Staubli VAL3: appLauncher.pjx

--- appLauncher.pjx ---
Parameters version=s8.21Cs9_BS4703 stackSize=200000 millimeterUnit=true
Program file=_getForce.pgx
Program file=_productCycle.pgx
Program file=_supervisorTasks.pgx
Program file=_systemStates.pgx
Program file=_tCycleCtrl.pgx
Program file=_TolleranceCheck.pgx
Program file=Init.pgx
Program file=kill.pgx
Program file=Main.pgx
Program file=search_traj.pgx
Program file=start.pgx
Program file=stop.pgx
Data file=appLauncher.dtx
Library alias=rs path=Disk://source/projectSource/robotStatus/robotStatus.pjx
Library alias=io path=Disk://source/projectSource/io/io.pjx
Library alias=home path=Disk://HMI_cs9/home/home.pjx
Library alias=plc path=Disk://source/projectSource/plc/plc.pjx
Library alias=prog path=Disk://source/projectSource/program/program.pjx
Library alias=program path=Disk://source/projectSource/program/program.pjx
Library alias=hmi_util path=Disk://HMI_cs9/HMI_util/HMI_util.pjx
Library alias=libTqe path=Disk://LibTorque/LibTorque.pjx
Library alias=trajectory path=Disk://source/projectSource/trajectory/trajectory.pjx
Library alias=ar path=Disk://autoReturn/autoReturn.pjx
Library alias=saveData path=Disk://source/saveData/saveData.pjx

--- appLauncher.dtx ---
bool _bAtHome
bool _bEndCycle
bool _bHeavyAlarm
bool _bIsScara
bool _bShowEndBt
bool _bShowPauseBt
bool _bShowResetBt
bool _bShowStartBt
bool _bShowStopBt
bool bBool
bool bControlByRobot = true
bool bTosave
frame test3 = {fatherId=world[0]}
num _nAvgCapacity
num _nBestCapacity
num _nCTIndex
num _nCapacity
num _nClock[10]
  [1] = 12488.271809
  [3] = 12488.271821
num _nCycleTime[10]
num _nLastStateCMD
num _nOmacStat
num _nStateCMD
num nCycleCmd
num nErrorCode = 1
num nLastLib
num nProgCode
string _sArmType
string _sOmacCmd
string _sOmacStatus = "1"
string _sPageAvergeCapacity
string _sPageBestCapacity
string _sPageCurrentCapacity
string _sPageCycleStatus
string _sPageHerej
string _sPagePosition
string _sPageProfile
string _sPageRobotStatus
string _sPageSN
string sMsg
num nForce[6]
public bool bGetMovId
mdesc mHome = {accel=20, vel=20, decel=20, blend=off}
string sSessionList
pointRx pPowerOFF = {fatherId=world[0]}
bool bMemState
pointRx pHere1 = {fatherId=world[0]}
pointRx pHere2 = {fatherId=world[0]}
bool bAutoConnectMove

--- Main.pgx ---
program Main()
  local bool l_bResult
  local bool l_bStartClock
  local num l_nClock
  local num l_nResult
begin
  //

  home:sVersion="version:5.0"
  resetMotion()
  //初始化
  //  call cycle_Init()
  //
  // userPage("StartUp")

  sMsg=">>> Loading 数据库 "+toString("",saveData:nLibIndex)+" <<<"
  //guohangxin add 2023.03.23
  //call initLib:initlib()
  saveData:nLibIndex=0
  call program:loadPROG(saveData:nLibIndex,l_nResult)
  call trajectory:loadTRAJ(saveData:nLibIndex,l_nResult)
  sMsg=""

  //机器人状态
  taskCreate "plc",60,plc:main()
  wait(taskStatus("plc")==1)
  //HMI
  taskCreate "HMI",50,home:main()
  wait(taskStatus("HMI")==1)
  //  //lifebit
  taskCreate "supervisorTask",10,_supervisorTasks()
  wait(taskStatus("supervisorTask")==1)
  do
    //机器人当前状态
    call _systemStates()
    //生产控制
    call _tCycleCtrl()
    //上下电位置记录
    // call _TolleranceCheck(bAutoConnectMove)
    delay(0)
  until rs:bQuitApp==true

  call kill()

end

--- start.pgx ---
program start()
begin
  taskCreate "appMain",100,Main()
end

--- _getForce.pgx ---
program _getForce()
  local num i
  local num l_nForce[6]
begin
  for i=0 to 5
    nForce[i]=0
  endFor

  do
    getJointForce(l_nForce)
    for i=0 to 5
      if abs(l_nForce[i])>nForce[i]
        nForce[i]=abs(l_nForce[i])
      endIf
    endFor
    //      if abs(l_nForce[4])>nForce[4]
    //        nForce[4]=abs(l_nForce[4])
    //      endIf
    //      if abs(l_nForce[5])>nForce[5]
    //        nForce[5]=abs(l_nForce[5])
    //      endIf
    delay(0)
  until rs:_nOmacStat==1
  //logMsg("程序号"+toString(".",rs:nProgCode)+"最大J5扭矩："+toString(".3",nForce[4])+",最大J6扭矩："+toString(".3",nForce[5]))
  rs:_sRobotStatus="程序号:"+toString(".",rs:nProgCode)+",J1MaxForce："+toString(".2",nForce[0])+",J2MaxForce："+toString(".2",nForce[1])+",J3MaxForce："+toString(".2",nForce[2])+",J4MaxForce："+toString(".2",nForce[3])+",J5MaxForce："+toString(".2",nForce[4])+",J6MaxForce："+toString(".2",nForce[5])
end

--- _productCycle.pgx ---
public program _productCycle()
  local bool l_bErr
  local bool l_bStartClock
  local num l_nClock
  local num l_nLastAct
  local num l_nLibIndex
  local string l_sPath
  local bool l_bFound
  local string l_sSelTraj
begin
  while true

    //
    //等待执行命令
    wait(plc:dInExcutePainting==true)
    //获取程序号
    call io:getAnaIO(io:aInItem[0].aAio,rs:nProgCode,l_bErr)
    //搜索对应traj
    call search_traj(l_bFound,l_sSelTraj,rs:nProgCode)
    //如果找到对应的traj，执行traj
    if l_bFound
      call trajectory:makeTraj(l_sSelTraj)
      waitEndMove()
    else
      popUpMsg("未找到喷涂号对应执行程序")
      rs:bIsError=true
      rs:bToStopCycle=true
    endIf
    delay(0)
  endWhile

  //  if l_bStartClock and l_nLastAct!=rs:nActCode
  //    rs:_nCTIndex=(rs:_nCTIndex+1)%size(rs:_nCycleTime)
  //    rs:_nCycleTime[rs:_nCTIndex]=clock()-l_nClock
  //  else
  //    l_bStartClock=true
  //  endIf
  //  l_nClock=clock()
  //  l_nLastAct=rs:nActCode
  //  //delay(0)
  //  //
  //  rs:_nOmacStat=1
  //  rs:sTrajStatus=""
  rs:_sRobotStatus="当前件生产结束"
  //2025.1.6 add 结束扭矩记录程序
  if taskStatus("getForce")!=-1
    delay(0.2)
    taskKill("getForce")
  endIf
end

--- _supervisorTasks.pgx ---
public program _supervisorTasks()
  local num l_i
  local bool l_bResult
begin
  for l_i = 0 to size(_nClock)-1
    _nClock[l_i]=0
  endFor
  do
    //任务监控
    if taskStatus("plc")>1 and (clock()-_nClock[1]>5)
      _nClock[1]=clock()
      taskResume("plc",0)
      rs:bIsError=true
    else
      _nClock[1]=clock()
    endIf
    if taskStatus("appMain")>1 and (clock()-_nClock[2]>5)
      _nClock[2]=clock()
      rs:bIsError=true
      taskResume("appMain",0)
    else
      _nClock[2]=clock()
    endIf
    if taskStatus("HMI")>1
      //保存当前数据
      bTosave=true
      call trajectory:onSave(bTosave)
      bTosave=true
      call program:onSave(bTosave)
      wait(rs:bIsSaving==false)
      l_bResult=userPageConfirm("需要重载HMI应用？")
      if l_bResult

        taskKill("HMI")
        wait(taskStatus("HMI")==-1)
        taskCreate "HMI",50,home:main()
        wait(taskStatus("HMI")==1)
      endIf
    endIf


    delay(0)
  until false
end

--- _systemStates.pgx ---
public program _systemStates()
begin
  // while true
  //程序运行中
  rs:bIsCycle=(taskStatus("cycle")>-1)
  //home
  rs:bIsHome=(abs(herej()-saveData:jHome)<{2,2,2,2,2,2})
  //使能上电
  rs:bPowerON=(isPowered()==true)
  //远程模式
  rs:bIsRemoteAuto=(workingMode()==4)
  //机器人正在移动
  rs:bIsMoving=(isSettled()==false)
  //机器人急停
  rs:bIsEstop=(esStatus()!=0)
  //
  rs:bIsReady=!rs:bIsCycle and rs:bIsHome and rs:bPowerON and !rs:bIsEstop and  rs:bIsRemoteAuto
  //程序报错
  rs:bIsError=(taskStatus("cycle")>1)

  // delay(0)
  // endWhile

end

--- _tCycleCtrl.pgx ---
program _tCycleCtrl()
  local bool l_bAckAlarm
  local bool l_bEndCmd
  local bool l_bErr
  local bool l_bHoldCmd
  local bool l_bPowerOff
  local bool l_bPowerOn
  local bool l_bResetCmd
  local bool l_bResetIO
  local bool l_bStartCmd
  local bool l_bStopCmd
  local num l_n
  local bool l_bResult
begin
  //启动程序
  if rs:bToStartCycle and rs:bIsReady
    rs:bToStartCycle=false
    taskCreate "cycle",100,_productCycle()
    wait(taskStatus("cycle")>-1)
  endIf
  //停止程序
  if(rs:bToStopCycle or rs:bIsEstop) and rs:bIsCycle
    rs:bToStopCycle=false
    resetMotion()
    stopMove()
    taskKill("cycle")
    wait(taskStatus("cycle")==-1)
  endIf
  //暂停程序
  if((rs:bToPause) and rs:bIsCycle) or taskStatus("cycle")>1
    rs:bToPause=false
    stopMove()
    rs:bIsPause=true
  endIf
  //暂停恢复程序
  if rs:bIsPause and rs:bIsCycle and rs:bToStartCycle
    rs:bToStartCycle=false
    rs:bIsPause=false
    if !isPowered()
      enablePower()
      l_bResult=watch(isPowered(),1)
      if !l_bResult
        logMsg("恢复生产任务上电超时")
        return
      endIf

    endIf
    autoConnectMove(true)
    restartMove()
  endIf
end

--- _TolleranceCheck.pgx ---
program _TolleranceCheck(bool& x_bAutoConnect)
  local string l_sMsg
begin

  if bMemState and !isPowered()
    pHere1=here(flange,world)
    l_sMsg="下电位置:"+toString(".2",pHere1.trsf.x)+","+toString(".2",pHere1.trsf.y)+","+toString(".2",pHere1.trsf.rz)
    logMsg(l_sMsg)
    bMemState=false
  elseIf !bMemState and isPowered()
    pHere2=here(flange,world)
    l_sMsg="上电位置:"+toString(".2",pHere1.trsf.x)+","+toString(".2",pHere1.trsf.y)+","+toString(".2",pHere1.trsf.rz)
    logMsg(l_sMsg)
    bMemState=true
  endIf
  //check
  if distance(pHere1.trsf,pHere2.trsf)<10
    x_bAutoConnect=true
  else
    x_bAutoConnect=false
    l_sMsg="TolleranceCheck位置偏差距离过大，需手动连接"
    popUpMsg(l_sMsg)
  endIf

end

--- Init.pgx ---
program Init()
  local num i
  local string l_sArmType
begin
  //dio

  //****************bool*****************
  _bEndCycle=false
  _bAtHome=false
  _bHeavyAlarm=false
  //判断是否是4轴机器人
  l_sArmType=left(getVersion("Arm Type"),2)
  _bIsScara=(l_sArmType=="rs" or l_sArmType=="ts" or l_sArmType=="tp")


  call rs:init()

end

--- kill.pgx ---
program kill()
begin
  //kill all task
  taskKill("safeCheck")
  taskKill("Reset")
  taskKill("Start")
  taskKill("Stop")
  taskKill("cycleCtrl")
  taskKill("plc")
  taskKill("lifebit")
  taskKill("actCtrl")
  taskKill("appMain")
  taskKill("HMI")

  //
  rs:bQuitApp=false
  stopMove()
  resetMotion()
  disablePower()
end

--- search_traj.pgx ---
program search_traj(bool& x_bFounded, string& x_sSessionName, num x_nSession)
  local string l_sEmpty
  local num i
  local num l_nSession
  local bool l_bOk
begin
  // init
  x_bFounded=false
  x_sSessionName=""
  //
  // get the list
  //
  l_sEmpty=""
  call trajectory:getTrajList(sSessionList)
  //
  // search the program from a number:
  //
  // "number+space+name"
  //
  // 01 MyPart
  // 10 YourPart
  //
  for i=0 to size(sSessionList)-1
    if sSessionList[i]!=""
      // convert the string "00 name" into a num
      toNum(sSessionList[i],l_nSession,l_bOk)
      if l_bOk and l_nSession==x_nSession
        x_sSessionName=sSessionList[i]
        x_bFounded=true
        // exit
        i=size(sSessionList)-1
      endIf
    endIf
  endFor
end

--- stop.pgx ---
program stop()
begin
  //kill all task
  taskKill("Reset")
  taskKill("Start")
  taskKill("Stop")
  taskKill("cycleCtrl")
  taskKill("Zones")
  taskKill("Main")
  taskKill("StatusRobot")
  //
  stopMove()
  resetMotion()
  disablePower()
end
